// Parameters of FB MON. Manual restart is active when the Restart port is connected.
TYPE
ST_SafeMonParameters :
STRUCT
    MonIn1MakeContact : BOOL;
    MonIn2MakeContact : BOOL;
    MonIn3MakeContact : BOOL;
    MonIn4MakeContact : BOOL;
    Secure1MakeContact : BOOL;
    Secure2MakeContact : BOOL;
    DiscrepancyTime1 : TIME; // MonIn1 / MonIn2
    DiscrepancyTime2 : TIME; // MonIn3 / MonIn4
    SecureDiscrepancyTime : TIME; // Secure1 / Secure2
    DelayTime : TIME; // switch-off delay of MonDelOut
    Edm1ResetTime : TIME;
    Edm2ResetTime : TIME;
    ManualFunctionTest : BOOL; // every connected MonIn pair must request the safe state once after start
    SafeInputsAfterDiscError : BOOL; // Safety Editor checkbox 'Safe Inputs after Disc Error', FALSE for a new block:
        // TRUE makes both channels of the pair that raised a discrepancy error return to the safe state together
        // before ErrAck can clear it
END_STRUCT
END_TYPE

(* stored: Version 1.1.0.1
   DUT ST_SafeMonParameters: Id {b7ad29f3-c8fa-5349-9b6f-af6e223c3780} *)
